// TIA Portal V19 export
// export: Created 2026-10-15T10:10:35.1362416Z, ExportSetting WithDefaults, DisplayName Totally Integrated Automation Portal, DisplayVersion V19, DisplayName TIA Portal Openness, DisplayVersion V19, DisplayName TIA Portal Version Control Interface, DisplayVersion V19, DisplayName STEP 7 Professional, DisplayVersion V19, DisplayName STEP 7 Safety, DisplayVersion V19, DisplayName WinCC Basic/Comfort/Advanced, DisplayVersion V19, DisplayName WinCC Unified, DisplayVersion V19
FUNCTION "ROLL_FB111" : Void   // FC13, SCL
{ S7_Optimized_Access := 'TRUE' }
VERSION : 0.1
// stored: AutoNumber true, IsIECCheckEnabled false, SetENOAutomatically false, UDAEnableTagReadback false
   VAR_TEMP
      preset : Word;
      signal : Bool;
   END_VAR
BEGIN

   #preset := W#16#2010;
   IF "ROLL_State".M[40, 5] THEN
       #preset := "ROLL_DB205".DW[5];
   ELSIF "ROLL_State".M[42, 1] THEN
       #preset := "ROLL_DB205".DW[17];
   ELSIF "ROLL_State".M[43, 5] THEN
       #preset := "ROLL_DB205".DW[25];
   ELSIF "ROLL_State".M[45, 2] THEN
       #preset := "ROLL_DB205".DW[33];
   END_IF;
   #signal := "ROLL_State".M[40, 5] OR "ROLL_State".M[42, 1] OR "ROLL_State".M[43, 5] OR "ROLL_State".M[45, 2]
   OR "ROLL_State".M[46, 5] OR "ROLL_State".M[48, 1] OR "ROLL_State".M[49, 5] OR "ROLL_State".M[51, 1];
   "ROLL_TimerOp"(Number := 1,
                  Operation := 0,
                  Signal := #signal,
                  Preset := #preset);
   IF (WORD_TO_INT("ROLL_TimerValue"(Number := 1)) <= 7)
       AND ("ROLL_State".M[40, 5] OR "ROLL_State".M[42, 1] OR "ROLL_State".M[43, 5]) AND "ROLL_State".M[111, 5] THEN
       "ROLL_State".M[58, 5] := TRUE;
   END_IF;
   IF "ROLL_State".M[63, 1] AND "ROLL_IO".Input[13, 3] THEN
       "ROLL_State".M[58, 5] := FALSE;
   END_IF;
   #preset := W#16#2010;
   IF "ROLL_State".M[41, 1] THEN
       #preset := "ROLL_DB205".DW[9];
   ELSIF "ROLL_State".M[42, 5] THEN
       #preset := "ROLL_DB205".DW[21];
   ELSIF "ROLL_State".M[44, 1] THEN
       #preset := "ROLL_DB205".DW[29];
   END_IF;
   #signal := "ROLL_State".M[41, 1] OR "ROLL_State".M[42, 5] OR "ROLL_State".M[44, 1]
   OR "ROLL_State".M[45, 6] OR "ROLL_State".M[47, 1] OR "ROLL_State".M[48, 5] OR "ROLL_State".M[50, 1];
   "ROLL_TimerOp"(Number := 2,
                  Operation := 0,
                  Signal := #signal,
                  Preset := #preset);
END_FUNCTION
